Fanuc KAREL source: KT00198.KL

PROGRAM KT00198
%NOLOCKGROUP
VAR
  B1: BOOLEAN
  Y2: ARRAY[2] OF BYTE
  OUT: INTEGER
BEGIN
  B1 = TRUE
    Y2[1] = 3
  OUT = B1 AND Y2[1]
END KT00198
